TYPE ST_DistanceCounter :
STRUCT
	lrAllOverDistance					:LREAL; 							(* All over counter distance *)
	lrAfterResetDistance				:LREAL; 							(* Counter distance since last reset *)
END_STRUCT
END_TYPE

(* stored: Version 1.1.0.1, ProductVersion 3.1.4024.15
   DUT ST_DistanceCounter: Id {c824c9cb-d929-4a9e-ad8c-836abed268fe} *)
